Fanuc KAREL source: KC00021.KL

PROGRAM KC00021
%NOLOCKGROUP
%ENVIRONMENT MOTN
VAR
  I: INTEGER
  J: INTEGER
  K: INTEGER
  R: REAL
  B: BOOLEAN
  S: STRING[80]
  T: STRING[80]
  P: PATH
  Q: PATH
  AI: ARRAY[8] OF INTEGER
  AB: ARRAY[244] OF BYTE
BEGIN
  B = MOTION_CTL
END KC00021
